Fanuc KAREL source: kt00733.KL

-- PROVISIONAL review KL for V1013-1; original PC SHA256 cd5244c12e56632da34401d4b07b44446b71641449ea9681d0666d7166a3627c
-- Incomplete behavior may be omitted. Consult companion uncertainty JSON. Do not deploy.
PROGRAM KT00733
%NOLOCKGROUP
VAR
  OUT : INTEGER
-- UNRESOLVED_DECL ARG type=002011
BEGIN
  -- UNRESOLVED_PC offsets 5-18; opcodes 22,1D,23
  -- UNRESOLVED_PC offsets 23-27; opcodes 7F
END KT00733
